Fanuc KAREL source: KB00025.KL

PROGRAM KB00025
%NOLOCKGROUP
%ENVIRONMENT IOSETUP
VAR
  P1: INTEGER
  P2: INTEGER
  P3: INTEGER
BEGIN
  P1 = 1
  P2 = 1
  P3 = 1
  CLR_PORT_SIM(P1, P2, P3)
END KB00025
